DATA_BLOCK "BlinkDb"
{ S7_Optimized_Access := 'TRUE' }
VERSION : 0.1
NON_RETAIN
"Blink"

BEGIN

END_DATA_BLOCK

